// TIA Portal V19 export
// export: Created 2026-10-15T10:10:36.3739301Z, ExportSetting WithDefaults, DisplayName Totally Integrated Automation Portal, DisplayVersion V19, DisplayName TIA Portal Openness, DisplayVersion V19, DisplayName TIA Portal Version Control Interface, DisplayVersion V19, DisplayName STEP 7 Professional, DisplayVersion V19, DisplayName STEP 7 Safety, DisplayVersion V19, DisplayName WinCC Basic/Comfort/Advanced, DisplayVersion V19, DisplayName WinCC Unified, DisplayVersion V19
FUNCTION "ROLL_PB17" : Void   // FC25, SCL
{ S7_Optimized_Access := 'TRUE' }
VERSION : 0.1
// stored: AutoNumber true, IsIECCheckEnabled false, SetENOAutomatically false, UDAEnableTagReadback false
   VAR_TEMP
      r : Bool;
      a1 : Word;
      a2 : Word;
      activeDataBlock : Int;
      comparisonResults : Array[0..0] of Bool;
   END_VAR
BEGIN

   #r := FALSE;
   #a1 := W#16#0000;
   #a2 := W#16#0000;
   #activeDataBlock := 0;
   // PB17, STEP 5 network 1
   #r := ((NOT "ROLL_State".M[70, 1]) AND "ROLL_State".M[3, 3]);
   "ROLL_State".M[70, 0] := #r;
   // PB17, STEP 5 network 2
   #r := "ROLL_State".M[70, 0];
   IF #r THEN
       "ROLL_State".M[70, 1] := TRUE;
   END_IF;
   #r := "ROLL_IO".Input[0, 2];
   IF #r THEN
       "ROLL_State".M[70, 1] := FALSE;
   END_IF;
   // PB17, STEP 5 network 3
   #r := ((("ROLL_IO".Input[0, 1] AND "ROLL_State".M[74, 1]) OR ("ROLL_IO".Input[0, 2] AND "ROLL_State".M[64, 0])) AND "ROLL_State".M[29, 1]);
   "ROLL_IO".Output[112, 0] := #r;
   // PB17, STEP 5 network 4
   #r := ((("ROLL_IO".Input[0, 1] AND "ROLL_State".M[74, 5]) OR ("ROLL_IO".Input[0, 2] AND "ROLL_State".M[64, 1])) AND "ROLL_State".M[29, 1]);
   "ROLL_IO".Output[112, 5] := #r;
   // PB17, STEP 5 network 5
   #r := (((("ROLL_IO".Input[0, 1] AND "ROLL_State".M[78, 4]) OR ("ROLL_IO".Input[0, 2] AND "ROLL_State".M[64, 4])) AND "ROLL_State".M[29, 0]) OR ("ROLL_IO".Output[113, 1] AND "ROLL_IO".Output[113, 3]));
   "ROLL_IO".Output[113, 1] := #r;
   // PB17, STEP 5 network 6
   #r := (((NOT "ROLL_State".M[71, 4]) AND "ROLL_State".M[71, 3]) OR ((("ROLL_IO".Input[0, 1] AND "ROLL_State".M[78, 6]) OR ("ROLL_IO".Input[0, 2] AND "ROLL_State".M[64, 5])) AND "ROLL_State".M[29, 0]));
   "ROLL_State".M[71, 3] := #r;
   // PB17, STEP 5 network 7
   #r := "ROLL_State".M[71, 3];
   "ROLL_IO".Output[113, 3] := #r;
   // PB17, STEP 5 network 8
   #r := (((NOT "ROLL_State".M[71, 3]) AND "ROLL_State".M[71, 4]) OR ((((NOT "ROLL_State".M[64, 5]) AND ((NOT "ROLL_State".M[20, 2]) OR "ROLL_IO".Input[124, 5]) AND "ROLL_IO".Input[0, 2]) OR ("ROLL_IO".Input[0, 1] AND "ROLL_State".M[78, 7])) AND "ROLL_State".M[29, 0]));
   "ROLL_State".M[71, 4] := #r;
   // PB17, STEP 5 network 9
   #r := "ROLL_State".M[71, 4];
   "ROLL_IO".Output[113, 2] := #r;
   // PB17, STEP 5 network 10
   #r := (("ROLL_IO".Input[0, 1] AND "ROLL_State".M[75, 4]) OR ("ROLL_IO".Input[0, 2] AND "ROLL_State".M[35, 2] AND "ROLL_State".M[65, 0]));
   "ROLL_State".M[79, 5] := #r;
   // PB17, STEP 5 network 11
   #r := ((NOT "ROLL_IO".Output[23, 0]) AND (NOT "ROLL_IO".Output[23, 4]) AND (NOT "ROLL_State".M[10, 3]) AND (NOT "ROLL_State".M[5, 0]) AND ((NOT "ROLL_IO".Input[11, 4]) OR (NOT "ROLL_IO".Input[11, 6])) AND "ROLL_IO".Input[11, 7] AND "ROLL_IO".Input[12, 5] AND "ROLL_IO".Input[12, 7] AND "ROLL_IO".Input[14, 0] AND "ROLL_State".M[29, 0] AND "ROLL_State".M[79, 5]);
   "ROLL_IO".Output[23, 1] := #r;
   // PB17, STEP 5 network 12
   #r := (("ROLL_IO".Input[0, 1] AND "ROLL_State".M[75, 5]) OR ("ROLL_IO".Input[0, 2] AND "ROLL_State".M[35, 2] AND "ROLL_State".M[65, 5]));
   "ROLL_State".M[79, 6] := #r;
   // PB17, STEP 5 network 13
   #r := ((NOT "ROLL_IO".Output[23, 1]) AND (NOT "ROLL_IO".Output[23, 4]) AND (NOT "ROLL_State".M[10, 2]) AND (NOT "ROLL_State".M[5, 0]) AND (((NOT "ROLL_IO".Input[119, 0]) AND "ROLL_State".M[0, 3]) OR (NOT "ROLL_IO".Input[11, 0]) OR (NOT "ROLL_IO".Input[11, 6])) AND "ROLL_IO".Input[11, 7] AND "ROLL_IO".Input[12, 5] AND "ROLL_IO".Input[12, 7] AND "ROLL_IO".Input[14, 0] AND "ROLL_State".M[29, 0] AND "ROLL_State".M[79, 6]);
   "ROLL_IO".Output[23, 0] := #r;
   // PB17, STEP 5 network 14
   #r := ((("ROLL_IO".Input[0, 1] AND "ROLL_State".M[75, 6]) OR ("ROLL_IO".Input[0, 2] AND "ROLL_State".M[35, 2] AND "ROLL_State".M[65, 6])) AND ("ROLL_IO".Output[23, 0] OR "ROLL_IO".Output[23, 1]));
   "ROLL_IO".Output[23, 3] := #r;
   // PB17, STEP 5 network 15
   #r := ((NOT "ROLL_IO".Output[23, 3]) AND ("ROLL_IO".Output[23, 0] OR "ROLL_IO".Output[23, 1]) AND ("ROLL_IO".Input[0, 1] OR "ROLL_State".M[31, 5]) AND "ROLL_State".M[29, 0]);
   "ROLL_IO".Output[23, 2] := #r;
   // PB17, STEP 5 network 16
   #r := (("ROLL_IO".Input[0, 1] AND "ROLL_State".M[76, 2]) OR ("ROLL_IO".Input[0, 2] AND "ROLL_State".M[35, 2] AND "ROLL_State".M[66, 4]));
   "ROLL_State".M[80, 0] := #r;
   // PB17, STEP 5 network 17
   #r := ((NOT "ROLL_IO".Output[23, 4]) AND (NOT "ROLL_State".M[10, 1]) AND (NOT "ROLL_State".M[5, 2]) AND (NOT "ROLL_State".M[9, 0]) AND ((NOT "ROLL_IO".Input[12, 5]) OR (NOT "ROLL_IO".Input[12, 7])) AND ("ROLL_IO".Input[124, 2] OR "ROLL_State".M[0, 4]) AND "ROLL_IO".Input[13, 0] AND "ROLL_IO".Input[13, 7] AND "ROLL_IO".Input[14, 0] AND "ROLL_State".M[29, 0] AND "ROLL_State".M[80, 0]);
   "ROLL_IO".Output[23, 5] := #r;
   // PB17, STEP 5 network 18
   #r := (("ROLL_IO".Input[0, 1] AND "ROLL_State".M[77, 0]) OR ("ROLL_IO".Input[0, 2] AND "ROLL_State".M[35, 2] AND "ROLL_State".M[66, 7]));
   "ROLL_State".M[80, 1] := #r;
   // PB17, STEP 5 network 19
   #r := "ROLL_IO".Input[12, 5];
   IF #r THEN
       "ROLL_State".M[80, 2] := TRUE;
   END_IF;
   #r := "ROLL_IO".Input[12, 1];
   IF #r THEN
       "ROLL_State".M[80, 2] := FALSE;
   END_IF;
   // PB17, STEP 5 network 20
   #r := (((("ROLL_IO".Input[11, 1] OR "ROLL_IO".Input[11, 2] OR "ROLL_IO".Input[11, 3] OR "ROLL_IO".Input[11, 4] OR "ROLL_IO".Input[119, 6] OR "ROLL_IO".Input[119, 7] OR "ROLL_IO".Input[120, 0] OR "ROLL_IO".Input[120, 1]) AND "ROLL_IO".Input[12, 1]) OR ("ROLL_IO".Input[11, 0] AND "ROLL_IO".Input[12, 1])) AND "ROLL_IO".Input[12, 7]);
   "ROLL_State".M[80, 6] := #r;
   // PB17, STEP 5 network 21
   #r := (("ROLL_IO".Input[11, 0] OR "ROLL_IO".Input[11, 1] OR "ROLL_IO".Input[11, 2] OR "ROLL_IO".Input[11, 3] OR "ROLL_IO".Input[11, 4] OR "ROLL_IO".Input[119, 6] OR "ROLL_IO".Input[119, 7] OR "ROLL_IO".Input[120, 0] OR "ROLL_IO".Input[120, 1]) AND "ROLL_IO".Input[12, 5] AND "ROLL_IO".Input[12, 7]);
   "ROLL_State".M[80, 7] := #r;
   // PB17, STEP 5 network 22
   #r := ((NOT "ROLL_IO".Output[23, 0]) AND (NOT "ROLL_IO".Output[23, 1]) AND (NOT "ROLL_IO".Output[23, 5]) AND (NOT "ROLL_State".M[10, 0]) AND (NOT "ROLL_State".M[5, 2]) AND (NOT "ROLL_State".M[80, 6]) AND ("ROLL_IO".Input[124, 2] OR "ROLL_State".M[0, 4]) AND "ROLL_IO".Input[13, 0] AND "ROLL_IO".Input[14, 0] AND "ROLL_State".M[29, 0] AND "ROLL_State".M[80, 1]);
   "ROLL_IO".Output[23, 4] := #r;
   // PB17, STEP 5 network 23
   #r := ((NOT "ROLL_State".M[68, 2]) AND (((NOT "ROLL_IO".Input[12, 5]) AND "ROLL_IO".Output[23, 5]) OR ("ROLL_IO".Output[23, 4] AND "ROLL_State".M[80, 2])));
   "ROLL_IO".Output[23, 7] := #r;
   // PB17, STEP 5 network 24
   #r := ((NOT "ROLL_IO".Output[23, 7]) AND ("ROLL_IO".Output[23, 4] OR "ROLL_IO".Output[23, 5]));
   "ROLL_IO".Output[23, 6] := #r;
   // PB17, STEP 5 network 25
   #r := (("ROLL_IO".Input[0, 1] AND "ROLL_State".M[77, 6]) OR ("ROLL_IO".Input[0, 2] AND "ROLL_State".M[35, 2] AND "ROLL_State".M[67, 0]));
   "ROLL_State".M[80, 3] := #r;
   // PB17, STEP 5 network 26
   #r := ((NOT "ROLL_IO".Output[112, 1]) AND (NOT "ROLL_IO".Output[113, 3]) AND (NOT "ROLL_IO".Input[124, 2]) AND (NOT "ROLL_State".M[10, 5]) AND (NOT "ROLL_State".M[70, 2]) AND (NOT "ROLL_State".M[9, 3]) AND "ROLL_IO".Input[11, 0] AND "ROLL_IO".Input[11, 6] AND "ROLL_IO".Input[12, 1] AND "ROLL_IO".Input[12, 7] AND "ROLL_State".M[29, 0] AND "ROLL_State".M[80, 3]);
   "ROLL_IO".Output[112, 2] := #r;
   // PB17, STEP 5 network 27
   #r := (("ROLL_IO".Input[0, 1] AND "ROLL_State".M[77, 4]) OR ("ROLL_IO".Input[0, 2] AND "ROLL_State".M[35, 2] AND "ROLL_State".M[67, 1]));
   "ROLL_State".M[80, 4] := #r;
   // PB17, STEP 5 network 28
   #r := ((NOT "ROLL_IO".Output[112, 2]) AND (NOT "ROLL_IO".Output[113, 3]) AND (NOT "ROLL_IO".Input[124, 1]) AND (NOT "ROLL_State".M[10, 4]) AND (NOT "ROLL_State".M[70, 2]) AND (NOT "ROLL_State".M[70, 3]) AND (NOT "ROLL_State".M[9, 3]) AND "ROLL_IO".Input[11, 0] AND "ROLL_IO".Input[11, 6] AND "ROLL_IO".Input[12, 1] AND "ROLL_IO".Input[12, 7] AND "ROLL_State".M[29, 0] AND "ROLL_State".M[80, 4]);
   "ROLL_IO".Output[112, 1] := #r;
   // PB17, STEP 5 network 29
   #r := ((("ROLL_IO".Input[0, 1] AND "ROLL_State".M[77, 7]) OR ("ROLL_IO".Input[0, 2] AND "ROLL_State".M[35, 2] AND "ROLL_State".M[67, 5])) AND "ROLL_State".M[29, 0]);
   "ROLL_IO".Output[112, 4] := #r;
   // PB17, STEP 5 network 30
   #r := ((("ROLL_IO".Input[0, 1] AND "ROLL_State".M[78, 0]) OR ("ROLL_IO".Input[0, 2] AND "ROLL_State".M[35, 2] AND "ROLL_State".M[67, 6])) AND "ROLL_State".M[29, 0]);
   "ROLL_IO".Output[112, 3] := #r;
   // PB17, STEP 5 network 31
   #r := ((NOT "ROLL_State".M[16, 0]) AND (NOT "ROLL_State".M[16, 1]) AND (NOT "ROLL_State".M[16, 2]) AND (NOT "ROLL_State".M[16, 4]) AND "ROLL_State".M[37, 2]);
   "ROLL_State".M[81, 4] := #r;
   // PB17, STEP 5 network 32
   RETURN;
END_FUNCTION
